SUBAPPLICATION GreenBlueBackground1_auxSC (* Hintergrundfarbe (TRUE -> Blau, FALSE -> Weiß) für 1 Objekt (Kompakt) *)
  (* Standard: 61499-2 *)
  (* Version 1.0, 2024-01-01, franz, Meisterschulen am Ostbahnhof *)
  PACKAGE MyLib::sys;
  IMPORT isobus::UT::Q::const::IDs::ID_NULL;
  IMPORT isobus::UT::Q::types::s1ObjectID;
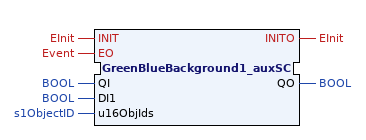
  EVENT_INPUT
    INIT : EInit; (* Initialization Request *)
    EO;
  END_EVENT
  EVENT_OUTPUT
    INITO : EInit; (* Initialization Confirm *)
  END_EVENT
  VAR_INPUT
    QI : BOOL := TRUE; (* Quality Input - TRUE to enable service *)
    DI1 : BOOL; (* Selector *)
    u16ObjIds : isobus::UT::Q::types::s1ObjectID := (u16ObjId := ID_NULL); (* Object IDs *)
  END_VAR
  VAR_OUTPUT
    QO : BOOL; (* Quality Output - TRUE if service executed successfully *)
  END_VAR
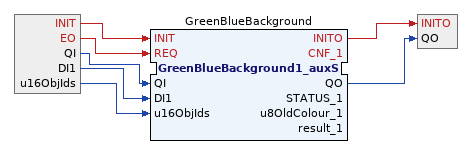
  SUBAPPS
    GreenBlueBackground : MyLib::sys::GreenBlueBackground1_auxS;
  END_SUBAPPS
  EVENT_CONNECTIONS
    EO TO GreenBlueBackground.REQ;
    INIT TO GreenBlueBackground.INIT;
    GreenBlueBackground.INITO TO INITO;
  END_CONNECTIONS
  DATA_CONNECTIONS
    u16ObjIds TO GreenBlueBackground.u16ObjIds;
    DI1 TO GreenBlueBackground.DI1;
    QI TO GreenBlueBackground.QI;
    GreenBlueBackground.QO TO QO;
  END_CONNECTIONS
END_SUBAPPLICATION
